Fanuc KAREL source: kd00004.KL

PROGRAM KD00004
%STACKSIZE=65535
%PRIORITY=65535
%NOLOCKGROUP
VAR
I : INTEGER
J : INTEGER
B : BOOLEAN
R : REAL
S : STRING[80]
BEGIN
I=1
END KD00004
